// TwinCAT 3 PLC project SendData
// ProgramVersion: 3.1.4023.0
// libraries:
//   Tc2_Standard, * (Beckhoff Automation GmbH)
//   Tc2_System, * (Beckhoff Automation GmbH)
//   Tc3_Module, * (Beckhoff Automation GmbH)
// project tree:
//   / PlcTask.TcTTO
//   POUs/ MAIN.TcPOU
// real-time tasks:
//   TASK PlcTask: cycle T#10ms, priority 20, ADS port 350
// I/O:
//   DEVICE Device 2 (EtherCAT), AmsNetId 192.168.18.191.3.1
//     Box 1 (sample_app) [sample_app]
// variable links:
//   SendData/SendData Instance <-> Device 2 (EtherCAT)/Box 1 (sample_app)
//     PlcTask Inputs/MAIN.rawAngle <-> Inputs process data mapping/Counter
//     PlcTask Outputs/MAIN.dummyData <-> Outputs process data mapping/Trigger

CONFIGURATION SendData
    RESOURCE PLC ON TwinCAT3
        TASK PlcTask(INTERVAL := T#10ms, PRIORITY := 20);
        PROGRAM MAIN WITH PlcTask : MAIN;
    END_RESOURCE
END_CONFIGURATION

// ---- POUs/MAIN.TcPOU
PROGRAM MAIN
VAR
	dir : BYTE := 1;
	speed : WORD := 100;
	dummyData AT %Q*: DWORD := SHL(dir,2*8) OR speed ;
	rawAngle AT %I*: DWORD;
	angle: REAL;
END_VAR

dummyData := SHL(dir,2*8) OR speed ;
angle := (rawAngle/100.0) - 180;

END_PROGRAM
